(* IEC 61131-3 sources: llm-plc-st-eval/codesys/dobles/A6, 10 files *)

(* ---- 01_Correcta.st ---- *)
(* DOBLE DE PRUEBA A6/Correcta - NO ES CORPUS. Esperado: veredicto 1 *)
FUNCTION_BLOCK FB_Modos
VAR_INPUT
    selector : INT;
    estadoSeguro : BOOL;
    cmdAuto : ARRAY[0..7] OF BOOL;
    cmdManual : ARRAY[0..7] OF BOOL;
    idxForzado : INT;
    valorForzado : BOOL;
    confirmarForzado : BOOL;
END_VAR
VAR_OUTPUT
    modoActivo : INT := 1;
    actuador : ARRAY[0..7] OF BOOL;
END_VAR
VAR
    forz : ARRAY[0..7] OF BOOL;
    prev : BOOL;
    flanco : BOOL;
    i : INT;
    selPrev : INT := 1;
END_VAR
IF estadoSeguro AND selector >= 0 AND selector <= 2 AND selector <> modoActivo THEN
    IF modoActivo = 2 THEN
        FOR i := 0 TO 7 DO
        forz[i] := FALSE;
    END_FOR
    END_IF
    modoActivo := selector;
END_IF
flanco := confirmarForzado AND NOT prev;
prev := confirmarForzado;
CASE modoActivo OF
    0:
        FOR i := 0 TO 7 DO
            actuador[i] := cmdAuto[i];
        END_FOR
    1:
        FOR i := 0 TO 7 DO
            actuador[i] := cmdManual[i];
        END_FOR
ELSE
    IF NOT estadoSeguro THEN
        FOR i := 0 TO 7 DO
        forz[i] := FALSE;
    END_FOR
    ELSIF flanco AND idxForzado >= 0 AND idxForzado <= 7 THEN
        forz[idxForzado] := valorForzado;
    END_IF
    FOR i := 0 TO 7 DO
        actuador[i] := forz[i];
    END_FOR
END_CASE
END_FUNCTION_BLOCK

(* ---- 02_ArrancaEnAuto.st ---- *)
(* DOBLE DE PRUEBA A6/ArrancaEnAuto - NO ES CORPUS. Esperado: veredicto 2, falla en el paso 0 *)
FUNCTION_BLOCK FB_Modos
VAR_INPUT
    selector : INT;
    estadoSeguro : BOOL;
    cmdAuto : ARRAY[0..7] OF BOOL;
    cmdManual : ARRAY[0..7] OF BOOL;
    idxForzado : INT;
    valorForzado : BOOL;
    confirmarForzado : BOOL;
END_VAR
VAR_OUTPUT
    modoActivo : INT := 0;
    actuador : ARRAY[0..7] OF BOOL;
END_VAR
VAR
    forz : ARRAY[0..7] OF BOOL;
    prev : BOOL;
    flanco : BOOL;
    i : INT;
    selPrev : INT := 1;
END_VAR
IF estadoSeguro AND selector >= 0 AND selector <= 2 AND selector <> modoActivo THEN
    IF modoActivo = 2 THEN
        FOR i := 0 TO 7 DO
        forz[i] := FALSE;
    END_FOR
    END_IF
    modoActivo := selector;
END_IF
flanco := confirmarForzado AND NOT prev;
prev := confirmarForzado;
CASE modoActivo OF
    0:
        FOR i := 0 TO 7 DO
            actuador[i] := cmdAuto[i];
        END_FOR
    1:
        FOR i := 0 TO 7 DO
            actuador[i] := cmdManual[i];
        END_FOR
ELSE
    IF NOT estadoSeguro THEN
        FOR i := 0 TO 7 DO
        forz[i] := FALSE;
    END_FOR
    ELSIF flanco AND idxForzado >= 0 AND idxForzado <= 7 THEN
        forz[idxForzado] := valorForzado;
    END_IF
    FOR i := 0 TO 7 DO
        actuador[i] := forz[i];
    END_FOR
END_CASE
END_FUNCTION_BLOCK

(* ---- 03_CambioSinSeguro.st ---- *)
(* DOBLE DE PRUEBA A6/CambioSinSeguro - NO ES CORPUS. Esperado: veredicto 2, falla en el paso 0 *)
FUNCTION_BLOCK FB_Modos
VAR_INPUT
    selector : INT;
    estadoSeguro : BOOL;
    cmdAuto : ARRAY[0..7] OF BOOL;
    cmdManual : ARRAY[0..7] OF BOOL;
    idxForzado : INT;
    valorForzado : BOOL;
    confirmarForzado : BOOL;
END_VAR
VAR_OUTPUT
    modoActivo : INT := 1;
    actuador : ARRAY[0..7] OF BOOL;
END_VAR
VAR
    forz : ARRAY[0..7] OF BOOL;
    prev : BOOL;
    flanco : BOOL;
    i : INT;
    selPrev : INT := 1;
END_VAR
IF selector >= 0 AND selector <= 2 AND selector <> modoActivo THEN
    IF modoActivo = 2 THEN
        FOR i := 0 TO 7 DO
        forz[i] := FALSE;
    END_FOR
    END_IF
    modoActivo := selector;
END_IF
flanco := confirmarForzado AND NOT prev;
prev := confirmarForzado;
CASE modoActivo OF
    0:
        FOR i := 0 TO 7 DO
            actuador[i] := cmdAuto[i];
        END_FOR
    1:
        FOR i := 0 TO 7 DO
            actuador[i] := cmdManual[i];
        END_FOR
ELSE
    IF NOT estadoSeguro THEN
        FOR i := 0 TO 7 DO
        forz[i] := FALSE;
    END_FOR
    ELSIF flanco AND idxForzado >= 0 AND idxForzado <= 7 THEN
        forz[idxForzado] := valorForzado;
    END_IF
    FOR i := 0 TO 7 DO
        actuador[i] := forz[i];
    END_FOR
END_CASE
END_FUNCTION_BLOCK

(* ---- 04_CambioSoloPorFlancoDeSelector.st ---- *)
(* DOBLE DE PRUEBA A6/CambioSoloPorFlancoDeSelector - NO ES CORPUS. Esperado: veredicto 2, falla en el paso 2 *)
FUNCTION_BLOCK FB_Modos
VAR_INPUT
    selector : INT;
    estadoSeguro : BOOL;
    cmdAuto : ARRAY[0..7] OF BOOL;
    cmdManual : ARRAY[0..7] OF BOOL;
    idxForzado : INT;
    valorForzado : BOOL;
    confirmarForzado : BOOL;
END_VAR
VAR_OUTPUT
    modoActivo : INT := 1;
    actuador : ARRAY[0..7] OF BOOL;
END_VAR
VAR
    forz : ARRAY[0..7] OF BOOL;
    prev : BOOL;
    flanco : BOOL;
    i : INT;
    selPrev : INT := 1;
END_VAR
IF selector <> selPrev AND estadoSeguro AND selector >= 0 AND selector <= 2 AND selector <> modoActivo THEN
    IF modoActivo = 2 THEN
        FOR i := 0 TO 7 DO
        forz[i] := FALSE;
    END_FOR
    END_IF
    modoActivo := selector;
END_IF
selPrev := selector;
flanco := confirmarForzado AND NOT prev;
prev := confirmarForzado;
CASE modoActivo OF
    0:
        FOR i := 0 TO 7 DO
            actuador[i] := cmdAuto[i];
        END_FOR
    1:
        FOR i := 0 TO 7 DO
            actuador[i] := cmdManual[i];
        END_FOR
ELSE
    IF NOT estadoSeguro THEN
        FOR i := 0 TO 7 DO
        forz[i] := FALSE;
    END_FOR
    ELSIF flanco AND idxForzado >= 0 AND idxForzado <= 7 THEN
        forz[idxForzado] := valorForzado;
    END_IF
    FOR i := 0 TO 7 DO
        actuador[i] := forz[i];
    END_FOR
END_CASE
END_FUNCTION_BLOCK

(* ---- 05_AceptaFueraDeRango.st ---- *)
(* DOBLE DE PRUEBA A6/AceptaFueraDeRango - NO ES CORPUS. Esperado: veredicto 2, falla en el paso 3 *)
FUNCTION_BLOCK FB_Modos
VAR_INPUT
    selector : INT;
    estadoSeguro : BOOL;
    cmdAuto : ARRAY[0..7] OF BOOL;
    cmdManual : ARRAY[0..7] OF BOOL;
    idxForzado : INT;
    valorForzado : BOOL;
    confirmarForzado : BOOL;
END_VAR
VAR_OUTPUT
    modoActivo : INT := 1;
    actuador : ARRAY[0..7] OF BOOL;
END_VAR
VAR
    forz : ARRAY[0..7] OF BOOL;
    prev : BOOL;
    flanco : BOOL;
    i : INT;
    selPrev : INT := 1;
END_VAR
IF estadoSeguro AND selector <> modoActivo THEN
    IF modoActivo = 2 THEN
        FOR i := 0 TO 7 DO
        forz[i] := FALSE;
    END_FOR
    END_IF
    modoActivo := selector;
END_IF
flanco := confirmarForzado AND NOT prev;
prev := confirmarForzado;
CASE modoActivo OF
    0:
        FOR i := 0 TO 7 DO
            actuador[i] := cmdAuto[i];
        END_FOR
    1:
        FOR i := 0 TO 7 DO
            actuador[i] := cmdManual[i];
        END_FOR
ELSE
    IF NOT estadoSeguro THEN
        FOR i := 0 TO 7 DO
        forz[i] := FALSE;
    END_FOR
    ELSIF flanco AND idxForzado >= 0 AND idxForzado <= 7 THEN
        forz[idxForzado] := valorForzado;
    END_IF
    FOR i := 0 TO 7 DO
        actuador[i] := forz[i];
    END_FOR
END_CASE
END_FUNCTION_BLOCK

(* ---- 06_MantenimientoSigueManual.st ---- *)
(* DOBLE DE PRUEBA A6/MantenimientoSigueManual - NO ES CORPUS. Esperado: veredicto 2, falla en el paso 6 *)
FUNCTION_BLOCK FB_Modos
VAR_INPUT
    selector : INT;
    estadoSeguro : BOOL;
    cmdAuto : ARRAY[0..7] OF BOOL;
    cmdManual : ARRAY[0..7] OF BOOL;
    idxForzado : INT;
    valorForzado : BOOL;
    confirmarForzado : BOOL;
END_VAR
VAR_OUTPUT
    modoActivo : INT := 1;
    actuador : ARRAY[0..7] OF BOOL;
END_VAR
VAR
    forz : ARRAY[0..7] OF BOOL;
    prev : BOOL;
    flanco : BOOL;
    i : INT;
    selPrev : INT := 1;
END_VAR
IF estadoSeguro AND selector >= 0 AND selector <= 2 AND selector <> modoActivo THEN
    IF modoActivo = 2 THEN
        FOR i := 0 TO 7 DO
        forz[i] := FALSE;
    END_FOR
    END_IF
    modoActivo := selector;
END_IF
flanco := confirmarForzado AND NOT prev;
prev := confirmarForzado;
CASE modoActivo OF
    0:
        FOR i := 0 TO 7 DO
            actuador[i] := cmdAuto[i];
        END_FOR
    1:
        FOR i := 0 TO 7 DO
            actuador[i] := cmdManual[i];
        END_FOR
ELSE
    IF NOT estadoSeguro THEN
        FOR i := 0 TO 7 DO
        forz[i] := FALSE;
    END_FOR
    ELSIF flanco AND idxForzado >= 0 AND idxForzado <= 7 THEN
        forz[idxForzado] := valorForzado;
    END_IF
    FOR i := 0 TO 7 DO
        actuador[i] := forz[i] OR cmdManual[i];
    END_FOR
END_CASE
END_FUNCTION_BLOCK

(* ---- 07_ForzadoNoRetiene.st ---- *)
(* DOBLE DE PRUEBA A6/ForzadoNoRetiene - NO ES CORPUS. Esperado: veredicto 2, falla en el paso 7 *)
FUNCTION_BLOCK FB_Modos
VAR_INPUT
    selector : INT;
    estadoSeguro : BOOL;
    cmdAuto : ARRAY[0..7] OF BOOL;
    cmdManual : ARRAY[0..7] OF BOOL;
    idxForzado : INT;
    valorForzado : BOOL;
    confirmarForzado : BOOL;
END_VAR
VAR_OUTPUT
    modoActivo : INT := 1;
    actuador : ARRAY[0..7] OF BOOL;
END_VAR
VAR
    forz : ARRAY[0..7] OF BOOL;
    prev : BOOL;
    flanco : BOOL;
    i : INT;
    selPrev : INT := 1;
END_VAR
IF estadoSeguro AND selector >= 0 AND selector <= 2 AND selector <> modoActivo THEN
    IF modoActivo = 2 THEN
        FOR i := 0 TO 7 DO
        forz[i] := FALSE;
    END_FOR
    END_IF
    modoActivo := selector;
END_IF
flanco := confirmarForzado AND NOT prev;
prev := confirmarForzado;
CASE modoActivo OF
    0:
        FOR i := 0 TO 7 DO
            actuador[i] := cmdAuto[i];
        END_FOR
    1:
        FOR i := 0 TO 7 DO
            actuador[i] := cmdManual[i];
        END_FOR
ELSE
    IF NOT estadoSeguro THEN
        FOR i := 0 TO 7 DO
        forz[i] := FALSE;
    END_FOR
    ELSIF flanco AND idxForzado >= 0 AND idxForzado <= 7 THEN
        forz[idxForzado] := valorForzado;
    END_IF
    FOR i := 0 TO 7 DO
        actuador[i] := forz[i];
    END_FOR
    IF NOT (flanco AND idxForzado >= 0 AND idxForzado <= 7) THEN
        FOR i := 0 TO 7 DO
        forz[i] := FALSE;
    END_FOR
    END_IF
END_CASE
END_FUNCTION_BLOCK

(* ---- 08_IdxSinValidar.st ---- *)
(* DOBLE DE PRUEBA A6/IdxSinValidar - NO ES CORPUS. Esperado: veredicto 2, falla en el paso 8 *)
FUNCTION_BLOCK FB_Modos
VAR_INPUT
    selector : INT;
    estadoSeguro : BOOL;
    cmdAuto : ARRAY[0..7] OF BOOL;
    cmdManual : ARRAY[0..7] OF BOOL;
    idxForzado : INT;
    valorForzado : BOOL;
    confirmarForzado : BOOL;
END_VAR
VAR_OUTPUT
    modoActivo : INT := 1;
    actuador : ARRAY[0..7] OF BOOL;
END_VAR
VAR
    forz : ARRAY[0..7] OF BOOL;
    prev : BOOL;
    flanco : BOOL;
    i : INT;
    selPrev : INT := 1;
END_VAR
IF estadoSeguro AND selector >= 0 AND selector <= 2 AND selector <> modoActivo THEN
    IF modoActivo = 2 THEN
        FOR i := 0 TO 7 DO
        forz[i] := FALSE;
    END_FOR
    END_IF
    modoActivo := selector;
END_IF
flanco := confirmarForzado AND NOT prev;
prev := confirmarForzado;
CASE modoActivo OF
    0:
        FOR i := 0 TO 7 DO
            actuador[i] := cmdAuto[i];
        END_FOR
    1:
        FOR i := 0 TO 7 DO
            actuador[i] := cmdManual[i];
        END_FOR
ELSE
    IF NOT estadoSeguro THEN
        FOR i := 0 TO 7 DO
        forz[i] := FALSE;
    END_FOR
    ELSIF flanco THEN
        forz[LIMIT(0, idxForzado, 7)] := valorForzado;
    END_IF
    FOR i := 0 TO 7 DO
        actuador[i] := forz[i];
    END_FOR
END_CASE
END_FUNCTION_BLOCK

(* ---- 09_SeguroNoAnula.st ---- *)
(* DOBLE DE PRUEBA A6/SeguroNoAnula - NO ES CORPUS. Esperado: veredicto 2, falla en el paso 11 *)
FUNCTION_BLOCK FB_Modos
VAR_INPUT
    selector : INT;
    estadoSeguro : BOOL;
    cmdAuto : ARRAY[0..7] OF BOOL;
    cmdManual : ARRAY[0..7] OF BOOL;
    idxForzado : INT;
    valorForzado : BOOL;
    confirmarForzado : BOOL;
END_VAR
VAR_OUTPUT
    modoActivo : INT := 1;
    actuador : ARRAY[0..7] OF BOOL;
END_VAR
VAR
    forz : ARRAY[0..7] OF BOOL;
    prev : BOOL;
    flanco : BOOL;
    i : INT;
    selPrev : INT := 1;
END_VAR
IF estadoSeguro AND selector >= 0 AND selector <= 2 AND selector <> modoActivo THEN
    IF modoActivo = 2 THEN
        FOR i := 0 TO 7 DO
        forz[i] := FALSE;
    END_FOR
    END_IF
    modoActivo := selector;
END_IF
flanco := confirmarForzado AND NOT prev;
prev := confirmarForzado;
CASE modoActivo OF
    0:
        FOR i := 0 TO 7 DO
            actuador[i] := cmdAuto[i];
        END_FOR
    1:
        FOR i := 0 TO 7 DO
            actuador[i] := cmdManual[i];
        END_FOR
ELSE
    IF flanco AND idxForzado >= 0 AND idxForzado <= 7 THEN
        forz[idxForzado] := valorForzado;
    END_IF
    FOR i := 0 TO 7 DO
        actuador[i] := forz[i];
    END_FOR
END_CASE
END_FUNCTION_BLOCK

(* ---- 10_SalirNoAnula.st ---- *)
(* DOBLE DE PRUEBA A6/SalirNoAnula - NO ES CORPUS. Esperado: veredicto 2, falla en el paso 15 *)
FUNCTION_BLOCK FB_Modos
VAR_INPUT
    selector : INT;
    estadoSeguro : BOOL;
    cmdAuto : ARRAY[0..7] OF BOOL;
    cmdManual : ARRAY[0..7] OF BOOL;
    idxForzado : INT;
    valorForzado : BOOL;
    confirmarForzado : BOOL;
END_VAR
VAR_OUTPUT
    modoActivo : INT := 1;
    actuador : ARRAY[0..7] OF BOOL;
END_VAR
VAR
    forz : ARRAY[0..7] OF BOOL;
    prev : BOOL;
    flanco : BOOL;
    i : INT;
    selPrev : INT := 1;
END_VAR
IF estadoSeguro AND selector >= 0 AND selector <= 2 AND selector <> modoActivo THEN
    modoActivo := selector;
END_IF
flanco := confirmarForzado AND NOT prev;
prev := confirmarForzado;
CASE modoActivo OF
    0:
        FOR i := 0 TO 7 DO
            actuador[i] := cmdAuto[i];
        END_FOR
    1:
        FOR i := 0 TO 7 DO
            actuador[i] := cmdManual[i];
        END_FOR
ELSE
    IF NOT estadoSeguro THEN
        FOR i := 0 TO 7 DO
        forz[i] := FALSE;
    END_FOR
    ELSIF flanco AND idxForzado >= 0 AND idxForzado <= 7 THEN
        forz[idxForzado] := valorForzado;
    END_IF
    FOR i := 0 TO 7 DO
        actuador[i] := forz[i];
    END_FOR
END_CASE
END_FUNCTION_BLOCK
